# EPICS substitutions: examples/PSI/best_practice/motion/stepper_bissc_hw_subst/cfg/hw.subs
#- ############################################################################
#- Master0
#-   0  0:0   PREOP  +  EK1100 EtherCAT-Koppler (2A E-Bus)
#-   1  0:1   PREOP  +  EL9227-5500 �berstromschutz 24V DC, 2K., max. 10A (Summe), eins
#-   2  0:2   PREOP  +  EL5042 2Ch. BiSS-C Encoder
#-   3  0:3   PREOP  +  EL5042 2Ch. BiSS-C Encoder
#-   4  0:4   PREOP  +  EL3204 4K. Ana. Eingang PT100 (RTD)
#-   5  0:5   PREOP  +  EL2008 8K. Dig. Ausgang 24V, 0.5A
#-   6  0:6   PREOP  +  EL1008 8K. Dig. Eingang 24V, 3ms
#-   7  0:7   PREOP  +  EL7041 1Ch. Stepper motor output stage (50V, 5A)
#-   8  0:8   PREOP  +  EL7041 1Ch. Stepper motor output stage (50V, 5A)
#-   9  0:9   PREOP  +  EL7041 1Ch. Stepper motor output stage (50V, 5A)
#-  10  0:10  PREOP  +  EL7041 1Ch. Stepper motor output stage (50V, 5A)

file "${ecmccomp_DIR}/HWTemplate.cmd" {
pattern { SLAVE_ID    HW_DESC       COMP                                COMP_CH   COMP_MACROS}

        { 0           EK1100        -1                                 -1         -1}
        { 1           EL9227-5500   -1                                 -1         -1}

# Encoders
        { 2           EL5042        Encoder-Renishaw-26bit-BISS-C       1         ""}
        { 2           EL5042        Encoder-Renishaw-26bit-BISS-C       2         ""}
        { 3           EL5042        -1                                 -1         -1}

# I/O
        {4            EL3204        -1                                 -1         -1}
        {5            EL2008        -1                                 -1         -1}
        {6            EL1008        -1                                 -1         -1}

# Drives
        {7            EL7041-0052   Motor-Generic-2Phase-Stepper        1         "I_MAX_MA=1000, I_STDBY_MA=500, U_NOM_MV=48000, R_COIL_MOHM=1230"}
        {8            EL7041-0052   Motor-Generic-2Phase-Stepper        1         "I_MAX_MA=1000, I_STDBY_MA=500, U_NOM_MV=48000, R_COIL_MOHM=1230"}
        {9            EL7041-0052   -1                                 -1         -1}
        {10           EL7041-0052   -1                                 -1         -1}
}
